(*
SPDX-FileCopyrightText: c 2026 Oleksandr Tiutyk <trofimich@gmail.com>
SPDX-License-Identifier: MIT
License: https://opensource.org/license/mit
*)

(*!
<summary>Checks scalar INT16 binding and positive and negative input values.</summary>
<description>
Uses a live case-owned automation parent and fresh local device fixtures on every run.
The scenario reads and writes ordinary simulated storage within one task cycle.
</description>
*)

{attribute 'no_assign'}
{attribute 'no_explicit_call' := 'do not call this function block directly'}
FUNCTION_BLOCK AnalogInputScalingAndScalarBindingTest EXTENDS TOF_Testing.SingleCycleTest
VAR_STAT
	{attribute 'hide'}
	_ClassName : STRING := __POUNAME();
END_VAR
VAR
	//! <summary>Live parent borrowed by the method-local simulated device.</summary>
	_AutomationRoot : MockAutomationController(name := "DevicesIORoot");
END_VAR

(*!
<summary>Checks scalar INT16 binding and positive and negative input values.</summary>
*)
METHOD PROTECTED ExecuteTest
VAR
	converter : TOF_Devices_IO.DirectAnalogValueConverter;
	analogInput : TOF_Devices_IO.AnalogInput(name := "AI_Scalar", parent := _AutomationRoot, converter := converter);
	rawInput : INT;
END_VAR
analogInput.Initialize();
analogInput.BindToInt16Value(rawValue := rawInput);

Assert.ThatBool(
	actual := analogInput.BoundToIO,
	message := "AnalogInput should be BoundToIO after BindToInt16Value"
).IsTrue();

rawInput := 5678;
analogInput.ProcessInput();

Assert.ThatLongReal(
	actual := analogInput.Value,
	message := "AnalogInput.Value should match raw INT input"
).ToBe(expected := 5678.0, tolerance := 0.001);

Assert.ThatBool(
	actual := analogInput.HasError,
	message := "AnalogInput should work without error when status is unbound"
).IsFalse();

rawInput := INT#-1234;
analogInput.ProcessInput();

Assert.ThatLongReal(
	actual := analogInput.Value,
	message := "Scalar input processing must preserve the INT16 sign"
).ToBe(expected := LREAL#-1234.0);
END_METHOD

//! <summary>Borrows the concrete class name. Callers must not modify it.</summary>
{attribute 'monitoring' := 'call'}
PROPERTY ClassName : REFERENCE TO STRING
GET
ClassName REF= _ClassName;
END_GET
END_PROPERTY

//! <summary>Borrows the compiler-initialized namespace name. Callers must not modify it.</summary>
{attribute 'monitoring' := 'call'}
PROPERTY NamespaceName : REFERENCE TO STRING
GET
NamespaceName REF= CurrentNamespace.Name;
END_GET
END_PROPERTY

//! <summary>Reports the concrete instance size in bytes.</summary>
{attribute 'monitoring' := 'call'}
PROPERTY SelfSize : ULINT
GET
SelfSize := XSIZEOF(THIS^);
END_GET
END_PROPERTY

END_FUNCTION_BLOCK

(* stored: Version 1.1.0.1
   POU AnalogInputScalingAndScalarBindingTest: Id {34e9d6aa-3a90-4250-824c-8a44f0e2cd93}, SpecialFunc None
   Method ExecuteTest: Id {83052bcc-187a-477e-986d-a457148425a5}
   Property ClassName: Id {6d73bd62-6bfa-49dc-ae6a-03b4cfa97410}
   Get Get: Id {5c0d7d75-74b5-4db8-bff2-adb943fe081a}
   Property NamespaceName: Id {1a5d5c9a-b753-401f-9e69-2b016e511fd2}
   Get Get: Id {949d7944-8be1-4cfd-989e-5e1812b83801}
   Property SelfSize: Id {af2b9357-3c7c-43aa-bd9a-8d625e28f0ca}
   Get Get: Id {8a9b890d-8a32-4944-aebb-3c5de5c1004b} *)
